Fanuc KAREL source: KD00057.KL

PROGRAM KD00057
%NOLOCKGROUP
%DEFGROUP = 1
VAR
  I: INTEGER
  J: INTEGER
  B: BOOLEAN
  R: REAL
  S: STRING[80]
  P: POSITION
  Q: POSITION
BEGIN
  MOVE TO P VIA Q
END KD00057
